// TIA Portal V21 export
// export: Created 2026-08-21T20:18:55.3555747Z, ExportSetting None, DisplayName Totally Integrated Automation Portal, DisplayVersion V21, DisplayName STEP 7 Professional, DisplayVersion V21, DisplayName STEP 7 Safety, DisplayVersion V21, DisplayName Tech WebApplication, DisplayVersion V21, DisplayName WinCC Basic/Comfort/Advanced, DisplayVersion V21, DisplayName WinCC Professional, DisplayVersion V21, DisplayName WinCC Unified, DisplayVersion V21
TYPE "UDT_MTP_ServiceControlExtended"
   STRUCT
      ServiceControl : "UDT_MTP_ServiceControl";
      ServiceSetup { S7_SetPoint := 'True'} : "UDT_Service_Setup";
   END_STRUCT;
END_TYPE
